SUBAPPLICATION Softkey_Aux_IXA_TO_Remote_WRITE_Option (* VT-SoftKey lesen ODER AUX-Zuweisung (Joystick) lesen ODER lokaler Web-Override (z.B. vt-ui-mirror auf demselben Modul) + Remote-OPC-UA-Write an Zielmodul (generisch, ein Kanal, ohne Status-Feedback) - Option-Lib-Variante von Softkey_Aux_IXA_TO_Remote_WRITE: alle 4 Bausteine mit eigenem QI (Softkey_IXA, Aux_IXA, SUBSCRIBE_WEB, AX_CLIENT_1_0) werden von einem einzigen Option::AOption-Socket sequenziell initialisiert und gated (echtes INIT_REQ/INIT_CNF statt bloss einem QI-Bool, Franz: 'muss ein AOption Adapter sein'). AOption_OUT reicht die Aktivierung an eine nachgeschaltete Gruppe weiter (Daisy-Chain, analog MyLib_AX_Option::sys::OptionalGroup_001a/Franz: 'ich zeige dir wie man 2 Dinge die zusammenhaengen machen kann') - fuer Softkey_Aux_IXA_TO_Remote_WRITE_BG_Option_OPC, wo die Status-Haelfte anschliessend dieselbe Option bekommt, und fuer mehrere SoftKeys, die dieselbe Option teilen (z.B. Bunker_Klappen_Auf -> Bunker_Klappen_Zu). *)
  (* Standard: 61499-2; Description: Copyright (c) 2026 Büngener Schuder GmbH This program and the accompanying materials are made available under the terms of the Eclipse Public License 2.0 which is available at https://www.eclipse.org/legal/epl-2.0/ SPDX-License-Identifier: EPL-2.0 *)
  (* Version 1.2, 2026-10-30, Franz Höpfinger, Büngener Schuder GmbH, Remote-Clients mit Remote_Init_Retry: Kette (und Option-INIT_CNF) wartet nicht mehr auf die Gegenstation, nach INITO- neuer Versuch nach 2 s (forte #1092, sonst 60 s pro fehlendem Node und danach tot). *)
  (* Version 1.1, 2026-10-13, Franz Höpfinger, Büngener Schuder GmbH, E_REND_3 (parallele Rendezvous-Variante) verworfen - Franz zeigte den etablierten Daisy-Chain-Stil (OptionalGroup_001a/b, training1): sequenzielle INIT-Verkettung (Softkey_IXA->Aux_IXA->SUBSCRIBE_WEB->AX_CLIENT_1_0) statt paralleler Rendezvous, plus neuer PLUG1-Ausgang (AOption_EVENT_TO_X) fuer Weiterverkettung. SUBSCRIBE_WEB jetzt auch gated (hat QI/INIT/INITO wie die anderen 3) - Franz: 'reicht es alle Bausteine auszumachen die einen QI haben'. *)
  (* Version 1.0, 2026-10-13, Franz Höpfinger, Büngener Schuder GmbH, initial implementation (verworfen, siehe v1.1) - Option-Lib-Variante von Softkey_Aux_IXA_TO_Remote_WRITE (bleibt fuer die 10+ nicht-optionalen Aufrufer unveraendert). *)
  PACKAGE MyLib::sys;
  IMPORT isobus::UT::Q::const::IDs::ID_NULL;
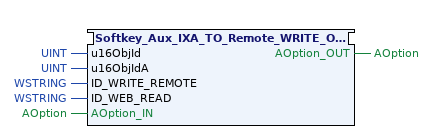
  VAR_INPUT
    u16ObjId : UINT := ID_NULL; (* Object ID SoftKey (VT) *)
    u16ObjIdA : UINT := ID_NULL; (* Object ID AuxFunction2 (VT) *)
    ID_WRITE_REMOTE : WSTRING; (* Remote-Write-Adresse zum Zielmodul (Befehl, ACTION=WRITE, CLIENT) *)
    ID_WEB_READ : WSTRING; (* Lokale Subscribe-Adresse fuer einen Web-Client (z.B. vt-ui-mirror) auf demselben Modul, ODER-verknuepft mit SoftKey und AUX *)
  END_VAR
  SOCKETS
    AOption_IN : Option::AOption; (* Treibt INIT/QI von Softkey_IXA/Aux_IXA/SUBSCRIBE_WEB/AX_CLIENT_1_0 - anschliessen an z.B. AOption_AUI_DEMUX_N.OUTx *)
  END_SOCKETS
  PLUGS
    AOption_OUT : Option::AOption; (* Reicht die Aktivierung an eine nachgeschaltete Gruppe weiter (Daisy-Chain) - unbenutzt lassen, wenn nichts weiter folgt *)
  END_PLUGS
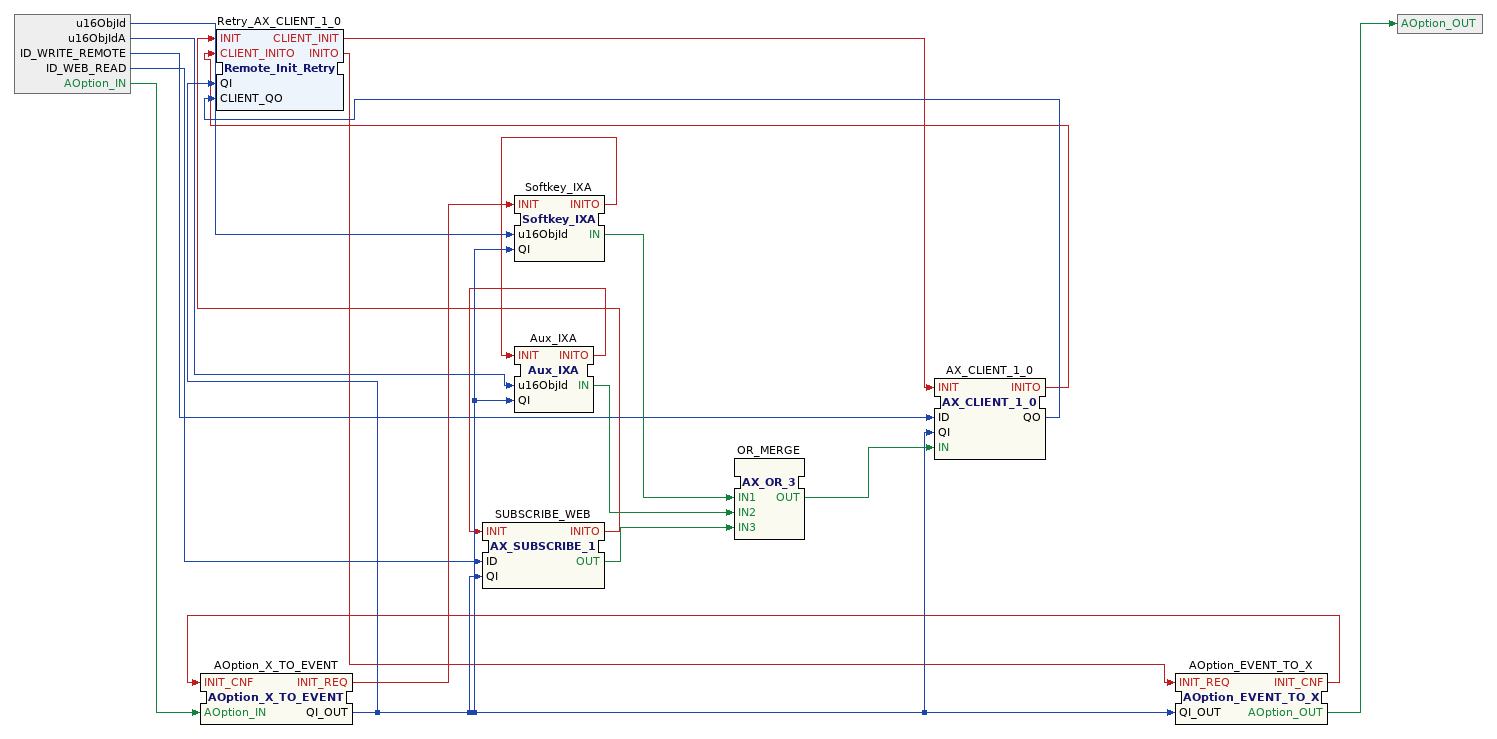
  FBS
    Softkey_IXA : isobus::UT::io::Softkey::Softkey_IXA;
    Aux_IXA : isobus::UT::io::Auxiliary::IN::Aux_IXA;
    SUBSCRIBE_WEB : adapter::net::AX_SUBSCRIBE_1;
    OR_MERGE : adapter::booleanOperators::AX_OR_3;
    AX_CLIENT_1_0 : adapter::net::AX_CLIENT_1_0;
    AOption_X_TO_EVENT : Option::conversion::AOption_X_TO_EVENT;
    AOption_EVENT_TO_X : Option::conversion::AOption_EVENT_TO_X;
  END_FBS
  SUBAPPS
    Retry_AX_CLIENT_1_0 : MyLib::sys::Remote_Init_Retry;
  END_SUBAPPS
  EVENT_CONNECTIONS
    SUBSCRIBE_WEB.INITO TO Retry_AX_CLIENT_1_0.INIT;
    Retry_AX_CLIENT_1_0.CLIENT_INIT TO AX_CLIENT_1_0.INIT;
    AX_CLIENT_1_0.INITO TO Retry_AX_CLIENT_1_0.CLIENT_INITO;
    Retry_AX_CLIENT_1_0.INITO TO AOption_EVENT_TO_X.INIT_REQ;
    AOption_X_TO_EVENT.INIT_REQ TO Softkey_IXA.INIT;
    Softkey_IXA.INITO TO Aux_IXA.INIT;
    Aux_IXA.INITO TO SUBSCRIBE_WEB.INIT;
    AOption_EVENT_TO_X.INIT_CNF TO AOption_X_TO_EVENT.INIT_CNF;
  END_CONNECTIONS
  DATA_CONNECTIONS
    AOption_X_TO_EVENT.QI_OUT TO Retry_AX_CLIENT_1_0.QI;
    AX_CLIENT_1_0.QO TO Retry_AX_CLIENT_1_0.CLIENT_QO;
    u16ObjId TO Softkey_IXA.u16ObjId;
    u16ObjIdA TO Aux_IXA.u16ObjId;
    ID_WEB_READ TO SUBSCRIBE_WEB.ID;
    ID_WRITE_REMOTE TO AX_CLIENT_1_0.ID;
    AOption_X_TO_EVENT.QI_OUT TO Softkey_IXA.QI;
    AOption_X_TO_EVENT.QI_OUT TO Aux_IXA.QI;
    AOption_X_TO_EVENT.QI_OUT TO SUBSCRIBE_WEB.QI;
    AOption_X_TO_EVENT.QI_OUT TO AX_CLIENT_1_0.QI;
    AOption_X_TO_EVENT.QI_OUT TO AOption_EVENT_TO_X.QI_OUT;
  END_CONNECTIONS
  ADAPTER_CONNECTIONS
    Softkey_IXA.IN TO OR_MERGE.IN1;
    Aux_IXA.IN TO OR_MERGE.IN2;
    SUBSCRIBE_WEB.OUT TO OR_MERGE.IN3;
    OR_MERGE.OUT TO AX_CLIENT_1_0.IN;
    AOption_IN TO AOption_X_TO_EVENT.AOption_IN;
    AOption_EVENT_TO_X.AOption_OUT TO AOption_OUT;
  END_CONNECTIONS
END_SUBAPPLICATION
